(*
SPDX-FileCopyrightText: © 2026 Oleksandr Tiutyk <trofimich@gmail.com>
SPDX-License-Identifier: MIT
License: https://opensource.org/license/mit
*)

(*!
<summary>Provides PLC execution context information and cached system time.</summary>
<description>
Task queries do not require Execute. A statically allocated TaskSystemState per cyclic PLC task owns its ADS
blocks and cached time. Execute and clock properties select the calling task. Outside cyclic context clock
getters return default values, SystemTime returns a null reference, and Execute and the interval setter do
nothing. Borrowed time references must not cross task boundaries.
</description>
*)

{attribute 'no_explicit_call' := 'do not call this function block directly'}
PROGRAM System
VAR CONSTANT
	(*!
	<summary>Number of entries in the generated PLC task information table.</summary>
	<description>
	Shared compile-time bound for per-task state arrays. Valid cyclic task indices range from 1 to TASK_COUNT;
	non-cyclic contexts are not entries.
	</description>
	*)
	TASK_COUNT : DINT := TO_DINT(XSIZEOF(TwinCAT_SystemInfoVarList._TaskInfo) / XSIZEOF(Global.PlcTaskSystemInfo));
END_VAR
VAR
	{attribute 'hide'}
	_ClassName : STRING := __POUNAME();

	{attribute 'hide'}
	_TaskStates : ARRAY [1..TASK_COUNT] OF TaskSystemState;
END_VAR

{attribute 'monitoring' := 'call'}
PROPERTY ClassName : REFERENCE TO STRING
GET
ClassName REF= _ClassName;
END_GET
END_PROPERTY

(*!
<summary>Converts calendar fields to a long date and time, preserving milliseconds.</summary>
<description>
The input must contain a valid date in the LDATE_AND_TIME range and milliseconds from 0 to 999. No timezone
conversion is performed.
</description>
*)

METHOD ConvertTimestructToLongDateTime : LDATE_AND_TIME
VAR_IN_OUT CONSTANT
	timestruct : Tc2_Utilities.TIMESTRUCT;
END_VAR
VAR
	longDateTimeLiteral : STRING;
END_VAR
longDateTimeLiteral := Strings.Concat255(
	'LDT#',
	TO_STRING(timestruct.wYear),
	'-',
	TO_STRING(timestruct.wMonth),
	'-',
	TO_STRING(timestruct.wDay),
	'-',
	TO_STRING(timestruct.wHour),
	':',
	TO_STRING(timestruct.wMinute),
	':',
	TO_STRING(timestruct.wSecond),
	'.',
	Tc2_Standard.RIGHT(STR := Tc2_Standard.CONCAT(STR1 := '00', STR2 := TO_STRING(timestruct.wMilliseconds)), SIZE := 3));
	
ConvertTimestructToLongDateTime := TO_LDT(longDateTimeLiteral);
END_METHOD

(*!
<summary>Advances system information requests and updates the cached clock.</summary>
<description>
Call cyclically from each task using system time. Advances only the calling task's ADS blocks and time
snapshot. Does nothing outside cyclic context. Read initial readiness through SystemDataValid; no result is
returned.
</description>
*)

METHOD Execute
VAR
	taskIndex : DINT;
END_VAR
taskIndex := GetCurrentTaskIndex();

IF taskIndex < 1 OR_ELSE taskIndex > TASK_COUNT THEN
	RETURN;
END_IF

_TaskStates[taskIndex].Execute();
END_METHOD

(*!
<summary>Borrows the runtime application information structure.</summary>
<description>
Returns a reference to TwinCAT_SystemInfoVarList._AppInfo. Treat runtime-owned information as read-only; the
call does not copy or refresh it.
</description>
*)
METHOD GetCurrentAppInfo : REFERENCE TO Global.PlcAppSystemInfo
GetCurrentAppInfo REF= TwinCAT_SystemInfoVarList._AppInfo;
END_METHOD

(*!
<summary>Identifies the calling execution context without accessing cached system data.</summary>
<description>
Returns a positive cyclic PLC task index, zero for a non-cyclic real-time context, or -1 for Windows context.
Does not allocate, log or raise exceptions and does not require Execute.
</description>
*)

METHOD PUBLIC GetCurrentTaskIndex : DINT
GetCurrentTaskIndex := Tc2_System.GETCURTASKINDEXEX();
END_METHOD

(*!
<summary>Returns a copy of the current cyclic PLC task information.</summary>
<description>
Does not require Execute. Outside a cyclic task, logs a diagnostic and returns default task information.
</description>
*)

METHOD GetCurrentTaskInfo : Global.PlcTaskSystemInfo
VAR
	taskIndex : DINT;
END_VAR
taskIndex := GetCurrentTaskIndex();

IF taskIndex > 0 THEN
	GetCurrentTaskInfo := TwinCAT_SystemInfoVarList._TaskInfo[taskIndex];
ELSE
	IF taskIndex < 0 THEN
		LogManager.TryLogMessage(
			message := "Method called from the Windows context",
			category := LOG_CATEGORY.ERROR,
			topic1 := TO_WSTRING(ClassName),
			topic2 := TO_WSTRING(__POUNAME())
		); 
	ELSE
		LogManager.TryLogMessage(
			message := "Method called not from a cyclic PLC task (such as FB_init)",
			category := LOG_CATEGORY.ERROR,
			topic1 := TO_WSTRING(ClassName),
			topic2 := TO_WSTRING(__POUNAME())
		); 
	END_IF
END_IF
END_METHOD

(*!
<summary>Returns the configured cycle duration of the calling cyclic PLC task.</summary>
<description>
Clears error on each call. Outside a cyclic task, returns zero and fills error without allocating an
exception. Does not require Execute. Outside cyclic context error timestamps are default values because there
is no task time snapshot.
</description>
*)

METHOD GetTaskCycleTime : LTIME
VAR_OUTPUT
	error : Error;
END_VAR
VAR
	taskInfo : Global.PlcTaskSystemInfo;
	taskIndex : DINT;
END_VAR
error.Clear();
taskIndex := GetCurrentTaskIndex();

IF taskIndex <= 0 THEN
	error.Fill(
		severity := ERROR_SEVERITY.ERROR,
		topSource := 'System.GetTaskCycleTime',
		rootSource := 'System.GetTaskCycleTime',
		topMessage := "Method requires a cyclic PLC task",
		rootMessage := "Method requires a cyclic PLC task",
		localTimestamp := SystemLocalDateTime,
		utcTimestamp := SystemUtcDateTime);
	GetTaskCycleTime := LTIME#0NS;
	RETURN;
END_IF

taskInfo := TwinCAT_SystemInfoVarList._TaskInfo[taskIndex];
GetTaskCycleTime := TO_LTIME(TO_ULINT(taskInfo.CycleTime) * ULINT#100);
END_METHOD

(*!
<summary>Returns the local AMS address obtained by the calling task.</summary>
<description>
Returns an empty address outside cyclic context or before acquisition. Address acquisition does not gate
SystemDataValid.
</description>
*)

PROPERTY FINAL LocalAmsNetId : Tc2_System.T_AmsNetID
GET
VAR
	taskIndex : DINT;
END_VAR
taskIndex := GetCurrentTaskIndex();

IF taskIndex < 1 OR_ELSE taskIndex > TASK_COUNT THEN
	RETURN;
END_IF

LocalAmsNetId := _TaskStates[taskIndex].LocalAmsNetId;
END_GET
END_PROPERTY

(*!
<summary>Provides the library namespace used in diagnostics.</summary>
<description>
Borrowed read-only reference to the compiler-initialized library namespace; no ownership transfer.
</description>
*)
{attribute 'monitoring' := 'call'}
PROPERTY NamespaceName : REFERENCE TO STRING
GET
NamespaceName REF= CurrentNamespace.Name;
END_GET
END_PROPERTY

(*!
<summary>Borrows the calling task's local calendar time for reading.</summary>
<description>
Returns a null reference outside cyclic context. In cyclic context the reference remains valid for the task
state lifetime, but its contents change on Execute. Read only after SystemDataValid; do not modify or share
this reference with another task.
</description>
*)

PROPERTY FINAL SystemTime : REFERENCE TO TIMESTRUCT
GET
VAR
	taskIndex : DINT;
END_VAR
SystemTime REF= 0;
taskIndex := GetCurrentTaskIndex();

IF taskIndex < 1 OR_ELSE taskIndex > TASK_COUNT THEN
	RETURN;
END_IF

SystemTime REF= _TaskStates[taskIndex].SystemTime;
END_GET
END_PROPERTY

(*!
<summary>Controls the calling task's clock synchronization interval in seconds.</summary>
<description>
Configure from the owning cyclic task using 1 to 86400 seconds. Each task has an independent interval. Outside
cyclic context the getter returns zero and the setter does nothing.
</description>
*)

PROPERTY FINAL SystemTimeSynchronisationInterval : DWORD
GET
VAR
	taskIndex : DINT;
END_VAR
taskIndex := GetCurrentTaskIndex();

IF taskIndex < 1 OR_ELSE taskIndex > TASK_COUNT THEN
	RETURN;
END_IF

SystemTimeSynchronisationInterval := _TaskStates[taskIndex].SystemTimeSynchronisationInterval;
END_GET
SET
VAR
	taskIndex : DINT;
END_VAR
taskIndex := GetCurrentTaskIndex();

IF taskIndex < 1 OR_ELSE taskIndex > TASK_COUNT THEN
	RETURN;
END_IF

_TaskStates[taskIndex].SystemTimeSynchronisationInterval := SystemTimeSynchronisationInterval;
END_SET
END_PROPERTY

(*!
<summary>Returns the calling task's cached timezone identifier.</summary>
<description>
Reads only the calling task's state without updating it. Returns the type's default value outside cyclic
context. Call Execute in this task and wait for SystemDataValid before consuming time values. Timezone
configuration is cached after initial acquisition of a known timezone; OS timezone configuration changes
require PLC application reinitialization.
</description>
*)

PROPERTY FINAL SystemTimeZoneId : Tc2_Utilities.E_TimeZoneID
GET
VAR
	taskIndex : DINT;
END_VAR
taskIndex := GetCurrentTaskIndex();

IF taskIndex < 1 OR_ELSE taskIndex > TASK_COUNT THEN
	RETURN;
END_IF

SystemTimeZoneId := _TaskStates[taskIndex].SystemTimeZoneId;
END_GET
END_PROPERTY

(*!
<summary>Returns a copy of the calling task's cached timezone rules.</summary>
<description>
Reads only the calling task's state without updating it. Returns the type's default value outside cyclic
context. Call Execute in this task and wait for SystemDataValid before consuming time values. Timezone
configuration is cached after initial acquisition of a known timezone; OS timezone configuration changes
require PLC application reinitialization.
</description>
*)

PROPERTY FINAL SystemTimeZoneInformation : Tc2_Utilities.ST_TimeZoneInformation
GET
VAR
	taskIndex : DINT;
END_VAR
taskIndex := GetCurrentTaskIndex();

IF taskIndex < 1 OR_ELSE taskIndex > TASK_COUNT THEN
	RETURN;
END_IF

SystemTimeZoneInformation := _TaskStates[taskIndex].SystemTimeZoneInformation;
END_GET
END_PROPERTY

(*!
<summary>Returns the local date and time captured by this task's last Execute.</summary>
<description>
Reads only the calling task's state without updating it. Returns the type's default value outside cyclic
context. Call Execute in this task and wait for SystemDataValid before consuming time values.
</description>
*)

PROPERTY FINAL SystemLocalDateTime : LDATE_AND_TIME
GET
VAR
	taskIndex : DINT;
END_VAR
taskIndex := GetCurrentTaskIndex();

IF taskIndex < 1 OR_ELSE taskIndex > TASK_COUNT THEN
	RETURN;
END_IF

SystemLocalDateTime := _TaskStates[taskIndex].SystemLocalDateTime;
END_GET
END_PROPERTY

(*!
<summary>Returns the UTC date and time captured by this task's last Execute.</summary>
<description>
Reads only the calling task's state without updating it. Returns the type's default value outside cyclic
context. Call Execute in this task and wait for SystemDataValid before consuming time values.
</description>
*)

PROPERTY FINAL SystemUtcDateTime : LDATE_AND_TIME
GET
VAR
	taskIndex : DINT;
END_VAR
taskIndex := GetCurrentTaskIndex();

IF taskIndex < 1 OR_ELSE taskIndex > TASK_COUNT THEN
	RETURN;
END_IF

SystemUtcDateTime := _TaskStates[taskIndex].SystemUtcDateTime;
END_GET
END_PROPERTY

(*!
<summary>Returns this task's cached local calendar time encoded as FILETIME.</summary>
<description>
Reads only the calling task's state without updating it. Returns the type's default value outside cyclic
context. Call Execute in this task and wait for SystemDataValid before consuming time values.
</description>
*)

PROPERTY FINAL SystemFileTime : Tc2_Utilities.T_FILETIME
GET
VAR
	taskIndex : DINT;
END_VAR
taskIndex := GetCurrentTaskIndex();

IF taskIndex < 1 OR_ELSE taskIndex > TASK_COUNT THEN
	RETURN;
END_IF

SystemFileTime := _TaskStates[taskIndex].SystemFileTime;
END_GET
END_PROPERTY

(*!
<summary>Returns this task's cached local calendar time encoded as 64-bit FILETIME.</summary>
<description>
Reads only the calling task's state without updating it. Returns the type's default value outside cyclic
context. Call Execute in this task and wait for SystemDataValid before consuming time values.
</description>
*)

PROPERTY FINAL SystemFileTime64 : Tc2_Utilities.T_FILETIME64
GET
VAR
	taskIndex : DINT;
END_VAR
taskIndex := GetCurrentTaskIndex();

IF taskIndex < 1 OR_ELSE taskIndex > TASK_COUNT THEN
	RETURN;
END_IF

SystemFileTime64 := _TaskStates[taskIndex].SystemFileTime64;
END_GET
END_PROPERTY

(*!
<summary>Indicates that the calling task has obtained system time and timezone successfully.</summary>
<description>
Latches initial time and timezone readiness for this task until application reinitialization. AMS Net ID does
not gate readiness. Returns FALSE outside cyclic context.
</description>
*)

PROPERTY FINAL SystemDataValid : BOOL
GET
VAR
	taskIndex : DINT;
END_VAR
taskIndex := GetCurrentTaskIndex();

IF taskIndex < 1 OR_ELSE taskIndex > TASK_COUNT THEN
	RETURN;
END_IF

SystemDataValid := _TaskStates[taskIndex].SystemDataValid;
END_GET
END_PROPERTY

END_PROGRAM

(* stored: Version 1.1.0.1
   POU System: Id {93357f84-3794-4f45-97d8-6aeeff54147a}, SpecialFunc None
   Folder Service methods: Id {cc1cd447-7df9-430c-b478-b2da6cfb4f5d}
   Property ClassName: Id {0f82d110-0834-4fc9-99f8-071cd51989f0}
   Get Get: Id {94979903-eeda-484e-add9-638420f45a0d}
   Method ConvertTimestructToLongDateTime: Id {c368065d-a4b5-46d7-baee-bf08cd6397d3}
   Method Execute: Id {0c6bf583-9275-4792-a0da-31f846086145}
   Method GetCurrentAppInfo: Id {972d2eff-4041-4c5b-bf4c-f1b03604e359}
   Method GetCurrentTaskIndex: Id {cc1072bd-3ddd-49d0-95e8-e9bd0e09202c}
   Method GetCurrentTaskInfo: Id {04f9a0b7-6093-424d-9fb3-0a09972c00e1}
   Method GetTaskCycleTime: Id {50bc18db-6507-4bea-bcbf-a26468abea5b}
   Property LocalAmsNetId: Id {f3ddb93d-d4f5-42d0-8950-99b61751e8a6}
   Get Get: Id {1d8d104b-6d8f-4619-bd22-ec259d3bad6c}
   Property NamespaceName: Id {33d380fa-ca9e-4f26-80e3-0dd39a24bf5e}
   Get Get: Id {c60ad75b-5af7-45b8-9e7c-d04b6018a6f3}
   Property SystemTime: Id {fc3dc1a5-f07a-44ea-8872-067f64602e6c}
   Get Get: Id {bca92c39-3456-4f53-b765-98dd8b8ca1e9}
   Property SystemTimeSynchronisationInterval: Id {e833856d-fead-4a01-a433-f36f3355afd1}
   Get Get: Id {ff6af129-621a-439f-9b9e-cfb3b139ccc1}
   Set Set: Id {88654d47-db1f-4874-a223-1856440fbe45}
   Property SystemTimeZoneId: Id {ab9dcc61-6d10-40c3-ac0d-cf0e93175250}
   Get Get: Id {16fd5c6a-37cb-4bf6-9aad-279fd5082ce8}
   Property SystemTimeZoneInformation: Id {b3056978-f770-4d50-b3df-5728e69da9eb}
   Get Get: Id {a946e3b2-b47c-4610-801d-30acfa22861c}
   Property SystemLocalDateTime: Id {d772a061-814f-43db-b63f-4c35be061290}
   Get Get: Id {4b089666-be80-48ce-a55b-c8a11b5d1f38}
   Property SystemUtcDateTime: Id {85aa966e-d1cf-4fc5-b00a-2bf21c99d4c1}
   Get Get: Id {b7db94d4-977e-4c63-a4db-2dfd7a348d17}
   Property SystemFileTime: Id {111195c9-20a9-426b-8d3b-6634564a7ce3}
   Get Get: Id {c8d3958a-6e2a-4a9e-9c2d-01d5f73efc76}
   Property SystemFileTime64: Id {82e61e7b-21eb-4a28-912e-f56fc8269f2e}
   Get Get: Id {1c7343e6-d74d-4e9e-bb43-a1f8ae551704}
   Property SystemDataValid: Id {0cb1ae30-8082-4885-a4df-b45f2a9ae686}
   Get Get: Id {b72f9f7c-20a1-4fe4-8dfb-5a17d0fca9a7} *)
